// TIA Portal V20 export
Screen "170Rollerup"  1276x673
  ScreenItem "permanentareaborderrectangle" at -1,0 size 0x0  Type=HmiRectangle
  ScreenItem "Line_Header_X0_Y64" at -1,65 size 1276x0  Type=HmiLine
  ScreenItem "Button_Back" at 1,2 size 90x60  Type=HmiButton
  ScreenItem "Title_ScreenOverview_X390_Y2_1" at 413,5 size 510x57  Type=HmiTextBox
  ScreenItem "Fusszeile_Button_ManualOPMode1_2" at 188,2 size 90x60  Type=HmiButton
  ScreenItem "Fusszeile_Button_ManualOPMode1_1" at 95,2 size 90x60  Type=HmiButton
  ScreenItem "Fusszeile_Button_ManualOPMode1_3" at 280,2 size 90x60  Type=HmiButton
  ScreenItem "Faceplate container_2" at 5,95 size 1270x134  Type=HmiFaceplateContainer
  ScreenItem "Move_Legend" at 1182,2 size 90x60  Type=HmiButton
  ScreenItem "文本域_3" at 1107,71 size 139x22  Type=HmiTextBox
  ScreenItem "面板容器_2" at 1090,4 size 88x58  Type=HmiFaceplateContainer
  ScreenItem "OPMode1_Blocked" at 1164,6 size 14x14  Type=HmiGraphicView
  ScreenItem "OPMode4_Foreground_Blocked" at 1092,5 size 88x58  Type=HmiGraphicView
